// LS Electric XG5000 project: NewProject
// PLC LSPLC
// module base 0 slot 0: 입력 모듈:XGI-D24A/B (DC 24V 입력, 32점 (전류소스 싱크공용/ 전류소스 입력))

PROGRAM NewProgram (task: 스캔 프로그램)

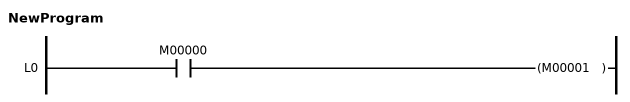
; L0
LOAD      M00000
OUT       M00001